(* IEC 61131-3 sources: IRIS-Project/LASAL CONTROL SOFTWARE/LasalProject_2025_09_12/Class/AutoManSelector, 1 file *)

(* ---- AutoManSelector.st ---- *)
(*!
<Class
	Name               = "AutoManSelector"
	Revision           = "0.0"
	RealtimeTask       = "false"
	CyclicTask         = "true"
	DefCyclictime      = "100 ms"
	BackgroundTask     = "false"
	Sigmatek           = "false"
	OSInterface        = "false"
	HighPriority       = "false"
	Automatic          = "false"
	UpdateMode         = "Prescan"
	SharedCommandTable = "true"
	Objectsize         = "(676,120)">
	<Channels>
		<Server Name="ClassSvr" Visualized="false" Initialize="false" WriteProtected="true" Retentive="false"/>
		<Server Name="s_EasyGUIEn" Visualized="false" Initialize="false" WriteProtected="false" Retentive="false"/>
		<Server Name="s_EmergencyStopMan" Visualized="false" Initialize="false" WriteProtected="false" Retentive="false"/>
		<Server Name="Selector" Visualized="false" Initialize="false" WriteProtected="false" Retentive="false"/>
		<Client Name="c_EasyGUIEn_IrrT" Required="true" Internal="false"/>
		<Client Name="c_EasyGUIEn_MainS" Required="true" Internal="false"/>
		<Client Name="ResetM1" Required="true" Internal="false"/>
		<Client Name="ResetM2" Required="true" Internal="false"/>
		<Client Name="ResetM3" Required="true" Internal="false"/>
		<Client Name="ResetM4" Required="true" Internal="false"/>
		<Client Name="ResetM5" Required="true" Internal="false"/>
		<Client Name="ResetM6" Required="true" Internal="false"/>
		<Client Name="ResetM7" Required="true" Internal="false"/>
		<Client Name="StopM1" Required="true" Internal="false"/>
		<Client Name="StopM2" Required="true" Internal="false"/>
		<Client Name="StopM3" Required="true" Internal="false"/>
		<Client Name="StopM4" Required="true" Internal="false"/>
		<Client Name="StopM5" Required="true" Internal="false"/>
		<Client Name="StopM6" Required="true" Internal="false"/>
		<Client Name="StopM7" Required="true" Internal="false"/>
		<Client Name="toAutomatic" Required="true" Internal="false"/>
		<Client Name="toManualM1" Required="true" Internal="false"/>
		<Client Name="toManualM2" Required="true" Internal="false"/>
		<Client Name="toManualM3" Required="true" Internal="false"/>
		<Client Name="toManualM4" Required="true" Internal="false"/>
		<Client Name="toManualM5" Required="true" Internal="false"/>
		<Client Name="toManualM6" Required="true" Internal="false"/>
		<Client Name="toManualM7" Required="true" Internal="false"/>
	</Channels>
	<Separators>
		<Clients>
			<SepChn Position="8"/>
			<SepChn Position="16"/>
			<SepChn Position="24"/>
		</Clients>
	</Separators>
</Class>
*)
AutoManSelector : CLASS
  //Servers:
	ClassSvr 	: SvrChCmd_DINT;
	Selector 	: SvrCh_DINT;
	s_EmergencyStopMan 	: SvrCh_DINT;
	s_EasyGUIEn 	: SvrCh_DINT;
  //Clients:
	toAutomatic 	: CltCh_DINT;
	toManualM1 	: CltCh_DINT;
	toManualM2 	: CltCh_DINT;
	toManualM3 	: CltCh_DINT;
	toManualM4 	: CltCh_DINT;
	toManualM5 	: CltCh_DINT;
	toManualM6 	: CltCh_DINT;
	toManualM7 	: CltCh_DINT;
	StopM1 	: CltCh_DINT;
	StopM2 	: CltCh_DINT;
	StopM3 	: CltCh_DINT;
	StopM4 	: CltCh_DINT;
	StopM5 	: CltCh_DINT;
	StopM6 	: CltCh_DINT;
	StopM7 	: CltCh_DINT;
	ResetM1 	: CltCh_DINT;
	ResetM2 	: CltCh_DINT;
	ResetM3 	: CltCh_DINT;
	ResetM4 	: CltCh_DINT;
	ResetM5 	: CltCh_DINT;
	ResetM6 	: CltCh_DINT;
	ResetM7 	: CltCh_DINT;
	c_EasyGUIEn_MainS 	: CltCh_DINT;
	c_EasyGUIEn_IrrT 	: CltCh_DINT;
  //Variables:
		v_Selector 	: DINT;
		v_EasyGUIEn 	: DINT;
  //Functions:

	FUNCTION VIRTUAL GLOBAL Init;

	FUNCTION VIRTUAL GLOBAL CyWork
		VAR_INPUT
			EAX 	: UDINT;
		END_VAR
		VAR_OUTPUT
			state (EAX) 	: UDINT;
		END_VAR;

	FUNCTION VIRTUAL GLOBAL Selector::Read
		VAR_OUTPUT
			output (EAX) 	: DINT;
		END_VAR;

	FUNCTION VIRTUAL GLOBAL s_EmergencyStopMan::Read
		VAR_OUTPUT
			output (EAX) 	: DINT;
		END_VAR;

	FUNCTION VIRTUAL GLOBAL s_EasyGUIEn::Read
		VAR_OUTPUT
			output (EAX) 	: DINT;
		END_VAR;
  //Tables:
	FUNCTION @STD
		VAR_OUTPUT
			ret_code	: CONFSTATES;
		END_VAR;
	FUNCTION GLOBAL TAB @CT_;
END_CLASS;

FUNCTION VIRTUAL GLOBAL AutoManSelector::Selector::Read
	VAR_OUTPUT
		output (EAX) 	: DINT;
	END_VAR

	output := Selector;

END_FUNCTION

FUNCTION VIRTUAL GLOBAL AutoManSelector::CyWork
	VAR_INPUT
		EAX 	: UDINT;
	END_VAR
	VAR_OUTPUT
		state (EAX) 	: UDINT;
	END_VAR

  v_Selector:=Selector.Read();
  v_EasyGUIEn:=s_EasyGUIEn.Read();

  if v_Selector=0 then
    toAutomatic.Write(input:=1);
    toManualM1.Write(input:=0);
    toManualM2.Write(input:=0);
    toManualM3.Write(input:=0);
    toManualM4.Write(input:=0);
    toManualM5.Write(input:=0);
    toManualM6.Write(input:=0);
    toManualM7.Write(input:=0);

  elsif v_Selector=1 then
    toAutomatic.Write(input:=0);
    toManualM1.Write(input:=1);
    toManualM2.Write(input:=1);
    toManualM3.Write(input:=1);
    toManualM4.Write(input:=1);
    toManualM5.Write(input:=1);
    toManualM6.Write(input:=1);
    toManualM7.Write(input:=1);

    case s_EmergencyStopMan of

    0:

    1:
      StopM1.Write(input:=1);
      StopM2.Write(input:=1);
      StopM3.Write(input:=1);
      StopM4.Write(input:=1);
      StopM5.Write(input:=1);
      StopM6.Write(input:=1);
      StopM7.Write(input:=1);
      s_EmergencyStopMan.Write(input:=2);

    2:
      StopM1.Write(input:=0);
      StopM2.Write(input:=0);
      StopM3.Write(input:=0);
      StopM4.Write(input:=0);
      StopM5.Write(input:=0);
      StopM6.Write(input:=0);
      StopM7.Write(input:=0);
      s_EmergencyStopMan.Write(input:=0);

    3:
      ResetM1.Write(input:=1);
      ResetM2.Write(input:=1);
      ResetM3.Write(input:=1);
      ResetM4.Write(input:=1);
      ResetM5.Write(input:=1);
      ResetM6.Write(input:=1);
      ResetM7.Write(input:=1);
      s_EmergencyStopMan.Write(input:=4);

    4:
      ResetM1.Write(input:=0);
      ResetM2.Write(input:=0);
      ResetM3.Write(input:=0);
      ResetM4.Write(input:=0);
      ResetM5.Write(input:=0);
      ResetM6.Write(input:=0);
      ResetM7.Write(input:=0);
      s_EmergencyStopMan.Write(input:=0);
    end_case;

  end_if;

  if v_EasyGUIEn then
    c_EasyGUIEn_MainS.Write(input:=1);
    c_EasyGUIEn_IrrT.Write(input:=1);
  else
    c_EasyGUIEn_MainS.Write(input:=0);
    c_EasyGUIEn_IrrT.Write(input:=0);
  end_if;

	state := READY;

END_FUNCTION

FUNCTION VIRTUAL GLOBAL AutoManSelector::Init

v_Selector:=0;
s_EasyGUIEn.Write(input:=1);
END_FUNCTION

FUNCTION VIRTUAL GLOBAL AutoManSelector::s_EmergencyStopMan::Read
	VAR_OUTPUT
		output (EAX) 	: DINT;
	END_VAR

	output := s_EmergencyStopMan;

END_FUNCTION

FUNCTION VIRTUAL GLOBAL AutoManSelector::s_EasyGUIEn::Read
	VAR_OUTPUT
		output (EAX) 	: DINT;
	END_VAR

	output := s_EasyGUIEn;

END_FUNCTION
